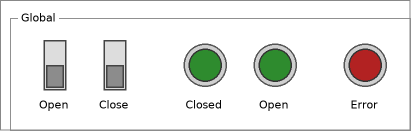
VISUALIZATION Cover  // 411x131
    GroupBox (10,10 401x121), "Global"
        DipSwitch (20,30 50x50), variable: MAIN.coverControl.bOpen, behaviour: TOGGLE, style: Switch-DipSwitch-Gray
        DipSwitch (80,30 50x50), variable: MAIN.coverControl.bClose, behaviour: TOGGLE, style: Switch-DipSwitch-Gray
        Lamp1 (170,30 50x50), variable: MAIN.coverControl.eCoverState = E_MirrorCoverState.closed, style: Lamp-Lamp1-Green
        Lamp1 (240,30 50x50), variable: MAIN.coverControl.eCoverState = E_MirrorCoverState.open, style: Lamp-Lamp1-Green
        Label (10,80 68x30), "Open"
        Label (70,80 68x30), "Close"
        Label (160,80 68x30), "Closed"
        Label (230,80 68x30), "Open"
        Lamp1 (330,30 50x50), variable: MAIN.coverControl.eCoverState = E_MirrorCoverState.error, style: Lamp-Lamp1-Red
        Label (320,80 68x30), "Error"
END_VISUALIZATION

(* stored: Version 1.1.0.1, ProductVersion 3.1.4024.15
   Visu Cover: Id {46ea3d6c-0d40-4863-8e54-1eda03fab11c} *)
